(* IEC 61131-3 sources: codesys-framework/txt/application/WeVe Utils (library)/TimeStamp/FB_TimeStampService/Feedback, 3 files *)

(* ---- TimeStamp_Local_AsString.prop.st ---- *)
PROPERTY TimeStamp_Local_AsString : STRING(23)

// --- BEGIN IMPLEMENTATION ---

// ----------- GET -----------
VAR
END_VAR

// -- BEGIN IMPLEMENTATION GET --
TimeStamp_Local_AsString := _sTimeStamp_Local_AsString;

(* ---- TimeStamp_UTC_AsString.prop.st ---- *)
PROPERTY TimeStamp_UTC_AsString : STRING(23)

// --- BEGIN IMPLEMENTATION ---

// ----------- GET -----------
VAR
END_VAR

// -- BEGIN IMPLEMENTATION GET --
TimeStamp_UTC_AsString := _sTimeStamp_UTC_AsString;

(* ---- TimeStampStringCreated.prop.st ---- *)
PROPERTY TimeStampStringCreated : BOOL

// --- BEGIN IMPLEMENTATION ---

// ----------- GET -----------
VAR
END_VAR

// -- BEGIN IMPLEMENTATION GET --
TimeStampStringCreated := _xTimeStampStringCreated;
